TYPE "DT_PAR_PID_CROSS_FLOW_VALVE_2"
VERSION : 0.1
   STRUCT
      INPUT_RAMP_MIN_VAL { S7_SetPoint := 'False'} : "DT_PARAM_SOLO" := (FALSE, 864, 0, 0.0, 0, T#0MS, 0.0, 0.0, '%');
      INPUT_RAMP_MAX_VAL { S7_SetPoint := 'False'} : "DT_PARAM_SOLO" := (FALSE, 865, 0, 0.0, 0, T#0MS, 0.0, 0.0, '%');
      INPUT_RAMP_FALLING_TIME { S7_SetPoint := 'False'} : "DT_PARAM_SOLO" := (FALSE, 866, 0, 0.0, 0, T#0MS, 0.0, 0.0, 's');
      INPUT_RAMP_RISING_TIME { S7_SetPoint := 'False'} : "DT_PARAM_SOLO" := (FALSE, 867, 0, 0.0, 0, T#0MS, 0.0, 0.0, 's');
      OUTPUT_RAMP_FALLING_TIME { S7_SetPoint := 'False'} : "DT_PARAM_SOLO" := (FALSE, 868, 0, 0.0, 0, T#0MS, 0.0, 0.0, 's');
      OUTPUT_RAMP_RISING_TIME { S7_SetPoint := 'False'} : "DT_PARAM_SOLO" := (FALSE, 869, 0, 0.0, 0, T#0MS, 0.0, 0.0, 's');
      MAN_ON { S7_SetPoint := 'False'} : "DT_PARAM_SOLO" := (FALSE, 870, 1, 0.0, 0, T#0MS, 0.0, 0.0, '-');
      P_SEL { S7_SetPoint := 'False'} : "DT_PARAM_SOLO" := (FALSE, 871, 1, 0.0, 0, T#0MS, 0.0, 0.0, '-');
      I_SEL { S7_SetPoint := 'False'} : "DT_PARAM_SOLO" := (FALSE, 872, 1, 0.0, 0, T#0MS, 0.0, 0.0, '-');
      INT_HOLD { S7_SetPoint := 'False'} : "DT_PARAM_SOLO" := (FALSE, 873, 1, 0.0, 0, T#0MS, 0.0, 0.0, '-');
      D_SEL { S7_SetPoint := 'False'} : "DT_PARAM_SOLO" := (FALSE, 874, 1, 0.0, 0, T#0MS, 0.0, 0.0, '-');
      NUM_OF_CYCLES { S7_SetPoint := 'False'} : "DT_PARAM_SOLO" := (FALSE, 875, 1, 0.0, 0, T#0MS, 0.0, 0.0, '-');
      GAIN { S7_SetPoint := 'False'} : "DT_PARAM_SOLO" := (FALSE, 876, 0, 0.0, 0, T#0MS, 0.0, 0.0, '');
      TI { S7_SetPoint := 'False'} : "DT_PARAM_SOLO" := (FALSE, 877, 1, 0.0, 0, T#0MS, 0.0, 0.0, '-');
      TD { S7_SetPoint := 'False'} : "DT_PARAM_SOLO" := (FALSE, 878, 1, 0.0, 0, T#0MS, 0.0, 0.0, '-');
      TM_LAG { S7_SetPoint := 'False'} : "DT_PARAM_SOLO" := (FALSE, 879, 1, 300.0, 0, T#0MS, 0.0, 0.0, '-');
      DEAD_W { S7_SetPoint := 'False'} : "DT_PARAM_SOLO" := (FALSE, 880, 0, 100.0, 0, T#0MS, 0.0, 0.0, '%');
      LMN_HLM { S7_SetPoint := 'False'} : "DT_PARAM_SOLO" := (FALSE, 881, 0, 30.0, 0, T#0MS, 0.0, 0.0, '%');
      LMN_LLM { S7_SetPoint := 'False'} : "DT_PARAM_SOLO" := (FALSE, 882, 0, 300.0, 0, T#0MS, 0.0, 0.0, '%');
      REF_MIN_VAL { S7_SetPoint := 'False'} : "DT_PARAM_SOLO" := (FALSE, 883, 0, 0.0, 0, T#0MS, 0.0, 0.0, '%');
      REF_MAX_VAL { S7_SetPoint := 'False'} : "DT_PARAM_SOLO" := (FALSE, 884, 0, 0.0, 0, T#0MS, 0.0, 0.0, '%');
      LMN_FAC { S7_SetPoint := 'False'} : "DT_PARAM_SOLO" := (FALSE, 885, 0, 0.0, 0, T#0MS, 0.0, 0.0, '-');
      LMN_OFFSET { S7_SetPoint := 'False'} : "DT_PARAM_SOLO" := (FALSE, 886, 0, 0.0, 0, T#0MS, 0.0, 0.0, '%');
      DISV { S7_SetPoint := 'False'} : "DT_PARAM_SOLO" := (FALSE, 887, 0, 0.0, 0, T#0MS, 0.0, 0.0, '-');
      MAN { S7_SetPoint := 'False'} : "DT_PARAM_SOLO" := (FALSE, 888, 0, 0.0, 0, T#0MS, 0.0, 0.0, '%');
      REFERENCE_CORRECTION { S7_SetPoint := 'False'} : "DT_PARAM_SOLO" := (FALSE, 889, 0, 0.0, 0, T#0MS, 0.0, 0.0, '-');
      OUT_CTRL_MODE { S7_SetPoint := 'False'} : "DT_PARAM_SOLO" := (FALSE, 890, 1, 0.0, 0, T#0MS, 0.0, 0.0, '-');
      SPARE_4 { S7_SetPoint := 'False'} : "DT_PARAM_SOLO" := (FALSE, 891, 0, 0.0, 0, T#0MS, 0.0, 0.0, '');
      SPARE_5 { S7_SetPoint := 'False'} : "DT_PARAM_SOLO" := (FALSE, 892, 0, 0.0, 0, T#0MS, 0.0, 0.0, '');
      SPARE_6 { S7_SetPoint := 'False'} : "DT_PARAM_SOLO" := (FALSE, 893, 0, 0.0, 0, T#0MS, 0.0, 0.0, '');
      SPARE_7 { S7_SetPoint := 'False'} : "DT_PARAM_SOLO" := (FALSE, 894, 0, 0.0, 0, T#0MS, 0.0, 0.0, '');
      SPARE_8 { S7_SetPoint := 'False'} : "DT_PARAM_SOLO" := (FALSE, 895, 0, 0.0, 0, T#0MS, 0.0, 0.0, '');
   END_STRUCT;

END_TYPE

